Fanuc KAREL source: KA00201.KL

PROGRAM KA00201
%NOLOCKGROUP
VAR
  SRC: ARRAY[4] OF VECTOR
  DST: ARRAY[4] OF BOOLEAN
BEGIN
  DST = SRC
END KA00201
